Fanuc KAREL source: kf00106.KL

-- PROVISIONAL review KL for V770-1; original PC SHA256 0f6864c519c97dc15ae682c627cfdf697c57f538b317bad0f9ca71ee23f068f6
-- Incomplete behavior may be omitted. Consult companion uncertainty JSON. Do not deploy.
PROGRAM KF00106
%NOLOCKGROUP
BEGIN
  -- UNRESOLVED_PC offsets 5-16; opcodes 2E,23
  -- UNRESOLVED_PC offsets 21-32; opcodes 2E,23
  -- UNRESOLVED_PC offsets 37-57; opcodes 27,27,9D,22,2A,22,31
  -- UNRESOLVED_PC offsets 62-66; opcodes 7F
END KF00106
